(*
	Span exporter test double. It keeps each accepted batch until the next one or free, and is
	busy while busy is set. callsWhileBusy counts export calls made while busy, which a processor
	must never make.
*)
FUNCTION_BLOCK FB_SpanExporter_ForInspection EXTENDS FB_SpanExporter_Base
VAR_INPUT
	busy: BOOL;
END_VAR
VAR_OUTPUT
	exportCount: UDINT;
	lastBatchCount: UDINT;
	tickCount: UDINT;
	callsWhileBusy: UDINT;
END_VAR

METHOD export : BOOL
VAR_IN_OUT
	spans: FB_SpanQueue;
END_VAR
VAR_INPUT
	count: UDINT;
END_VAR
VAR_OUTPUT
	failureReason: E_SpanExporterFailureReason;
END_VAR
IF THIS^.isBusy() THEN
	THIS^.callsWhileBusy := THIS^.callsWhileBusy + 1;
END_IF
export := SUPER^.export(spans:=spans, count:=count, failureReason=>failureReason);
IF export THEN
	THIS^.exportCount := THIS^.exportCount + 1;
	THIS^.lastBatchCount := THIS^._spans.count;
	// nothing is delivered, so the batch stays held until the next one or free
	THIS^._exportActive := FALSE;
END_IF
END_METHOD

(* The oldest span of the held batch, borrowed; 0 when nothing is held. *)
METHOD heldSpan : POINTER TO FB_Span
THIS^._spans.reset();
heldSpan := THIS^._spans.next();
END_METHOD

METHOD isBusy : BOOL
isBusy := THIS^.busy;
END_METHOD

METHOD tick : BOOL
VAR_OUTPUT
	failureReason: E_SpanExporterFailureReason;
END_VAR
THIS^.tickCount := THIS^.tickCount + 1;
failureReason := E_SpanExporterFailureReason.NA;
tick := TRUE;
END_METHOD

END_FUNCTION_BLOCK

(* stored: Version 1.1.0.1
   POU FB_SpanExporter_ForInspection: Id {d1e2c112-170e-4b6c-a2ea-96eff9a8f2f0}, SpecialFunc None
   Method export: Id {bfc15f05-cec6-465d-b91d-85232c0b1e2a}
   Method heldSpan: Id {9722e731-cc23-454b-a111-6ad1d8c6dad6}
   Method isBusy: Id {e6675821-044b-4c3e-a7d6-fced08703e57}
   Method tick: Id {62360fd4-efc1-479a-9eda-9e94368503c5} *)
